Fanuc KAREL source: kx00012.KL

-- PROVISIONAL review KL for V770-1; original PC SHA256 9a2d03ae288d398bedba258e9b741621f8630a5a6ac05282fcc9739969b625ef
-- Incomplete behavior may be omitted. Consult companion uncertainty JSON. Do not deploy.
PROGRAM KX00012
%NOLOCKGROUP
VAR
  I : INTEGER
  J : INTEGER
  B : BOOLEAN
  F : FILE
  S : STRING[80]
-- UNRESOLVED_DECL P type=000102
BEGIN
  -- UNRESOLVED_PC offsets 5-7; opcodes 9C,66
  -- UNRESOLVED_PC offsets 12-16; opcodes 7F
END KX00012
